Fanuc KAREL source: kb00177.KL

-- PROVISIONAL review KL for V1013-1; original PC SHA256 6897bbe3f41a19e3562888b8a6547c04313cf37196574e20eb8cb8e3a93b3ce4
-- Incomplete behavior may be omitted. Consult companion uncertainty JSON. Do not deploy.
PROGRAM KB00177
%NOLOCKGROUP
BEGIN
  -- UNRESOLVED_PC offsets 5-12; opcodes 9D,23
  -- UNRESOLVED_PC offsets 17-24; opcodes 9D,23
  -- UNRESOLVED_PC offsets 29-44; opcodes 2E,22,32,35
  -- UNRESOLVED_PC offsets 49-56; opcodes 9D,23
  -- UNRESOLVED_PC offsets 61-97; opcodes 27,22,22,22,1C,22,27,9D,31
  -- UNRESOLVED_PC offsets 102-106; opcodes 7F
END KB00177
